(* IEC 61131-3 sources: llm-plc-st-eval/data/definitivo/gemini-3.1-pro-preview/C4/few_shot, 3 files *)

(* ---- ejec_1.st ---- *)
El bloque de función `FB_D` implementa un sistema de control de alternancia y respaldo para dos bombas (sistema de trabajo-reserva o *duty-standby*). Cada vez que se recibe una nueva señal de demanda, el bloque alterna el turno de la bomba principal para garantizar un desgaste uniforme de ambos equipos. Durante la demanda, si la bomba a la que le corresponde el turno presenta una falla, el sistema activa automáticamente la bomba de respaldo y enciende una alarma. Cuando la demanda desaparece, ambas bombas y la alarma se apagan. Esta lógica es ideal para aplicaciones de bombeo de agua, sistemas de presión constante, estaciones de cárcamo, compresores o sistemas de lubricación redundantes donde la fiabilidad y el uso equilibrado de los motores son críticos.

```iecst
FUNCTION_BLOCK FB_D
VAR_INPUT
    demanda : BOOL; (* Señal de peticion de arranque del sistema *)
    falla1 : BOOL;  (* Señal de falla de la bomba 1 *)
    falla2 : BOOL;  (* Señal de falla de la bomba 2 *)
END_VAR
VAR_OUTPUT
    bomba1 : BOOL;   (* Comando de activacion para la bomba 1 *)
    bomba2 : BOOL;   (* Comando de activacion para la bomba 2 *)
    almFalla : BOOL; (* Alarma de falla en la bomba titular del turno *)
END_VAR
VAR
    turno : BOOL;    (* Bandera para alternar el turno (TRUE = Bomba 1, FALSE = Bomba 2) *)
    fDem : R_TRIG;   (* Detector de flanco de subida para la señal de demanda *)
END_VAR

(* Deteccion del flanco de subida de la señal de demanda *)
fDem(CLK := demanda);

(* Alternancia de turno con cada nueva demanda para equilibrar el desgaste *)
IF fDem.Q THEN
    turno := NOT turno;
END_IF

(* Logica de control de bombas mientras exista demanda *)
IF demanda THEN
    IF turno THEN
        (* Turno de la bomba 1 como principal *)
        bomba1 := NOT falla1;            (* Enciende bomba 1 si no tiene falla *)
        bomba2 := falla1 AND NOT falla2; (* Respaldo: enciende bomba 2 si la 1 falla y la 2 esta disponible *)
        almFalla := falla1;              (* Activa alarma si la bomba titular (1) falla *)
    ELSE
        (* Turno de la bomba 2 como principal *)
        bomba2 := NOT falla2;            (* Enciende bomba 2 si no tiene falla *)
        bomba1 := falla2 AND NOT falla1; (* Respaldo: enciende bomba 1 si la 2 falla y la 1 esta disponible *)
        almFalla := falla2;              (* Activa alarma si la bomba titular (2) falla *)
    END_IF
ELSE
    (* Apagado general del sistema cuando no hay demanda *)
    bomba1 := FALSE;
    bomba2 := FALSE;
    almFalla := FALSE;
END_IF
END_FUNCTION_BLOCK
```

(* ---- ejec_2.st ---- *)
Este bloque de función (FB_D) controla un sistema redundante de dos bombas con alternancia automática y lógica de respaldo (failover). Cada vez que se recibe una nueva señal de demanda, el sistema alterna el "turno" de la bomba principal para garantizar un desgaste equitativo entre ambas. Si la bomba a la que le corresponde el turno presenta una falla, el bloque arranca automáticamente la bomba de respaldo (siempre que esta no esté en falla también) y activa una alarma. Cuando la demanda desaparece, ambas bombas y la alarma se apagan. Esta lógica es ideal para aplicaciones de alta disponibilidad como estaciones de bombeo de agua potable, sistemas de achique (cárcamos), o circuitos de refrigeración/calefacción (HVAC) donde se requiere rotación de equipos y seguridad ante fallos.

```iecst
FUNCTION_BLOCK FB_D
VAR_INPUT
    demanda : BOOL; (* Señal de peticion de arranque del sistema *)
    falla1 : BOOL;  (* Señal de falla de la bomba 1 *)
    falla2 : BOOL;  (* Señal de falla de la bomba 2 *)
END_VAR
VAR_OUTPUT
    bomba1 : BOOL;   (* Comando de arranque para la bomba 1 *)
    bomba2 : BOOL;   (* Comando de arranque para la bomba 2 *)
    almFalla : BOOL; (* Alarma de falla de la bomba en turno *)
END_VAR
VAR
    turno : BOOL;    (* Memoria de alternancia (TRUE = Bomba 1, FALSE = Bomba 2) *)
    fDem : R_TRIG;   (* Detector de flanco de subida para la señal de demanda *)
END_VAR

(* Deteccion del flanco de subida de la demanda *)
fDem(CLK := demanda);

(* Alternancia del turno de la bomba principal en cada nueva demanda *)
IF fDem.Q THEN
    turno := NOT turno;
END_IF

(* Logica de control mientras la demanda este activa *)
IF demanda THEN
    IF turno THEN
        (* Turno de la bomba 1 como principal *)
        bomba1 := NOT falla1;                    (* Arranca bomba 1 si no tiene falla *)
        bomba2 := falla1 AND NOT falla2;         (* Respaldo: arranca bomba 2 si la 1 falla y la 2 esta disponible *)
        almFalla := falla1;                      (* Activa alarma si la bomba principal del turno fallo *)
    ELSE
        (* Turno de la bomba 2 como principal *)
        bomba2 := NOT falla2;                    (* Arranca bomba 2 si no tiene falla *)
        bomba1 := falla2 AND NOT falla1;         (* Respaldo: arranca bomba 1 si la 2 falla y la 1 esta disponible *)
        almFalla := falla2;                      (* Activa alarma si la bomba principal del turno fallo *)
    END_IF
ELSE
    (* Si no hay demanda, se apagan las bombas y la alarma *)
    bomba1 := FALSE;
    bomba2 := FALSE;
    almFalla := FALSE;
END_IF
END_FUNCTION_BLOCK
```

(* ---- ejec_3.st ---- *)
Este bloque de función (FB_D) controla un sistema redundante de dos bombas con alternancia automática y respaldo por falla. Cada vez que se recibe una nueva señal de demanda, el sistema alterna el "turno" de la bomba titular para equilibrar el desgaste mecánico de ambos equipos. Durante la operación, si la bomba que tiene el turno presenta una falla, el sistema activa automáticamente la bomba de respaldo (siempre y cuando esta no tenga falla también) y emite una alarma. Cuando no hay demanda, ambas bombas y la alarma se apagan. Es una aplicación clásica y muy útil para estaciones de bombeo de agua, sistemas de achique, circuitos de refrigeración o sistemas de lubricación donde se requiere alta disponibilidad y desgaste uniforme.

```iecst
FUNCTION_BLOCK FB_D
VAR_INPUT
    demanda : BOOL; (* Señal de peticion de arranque del sistema *)
    falla1 : BOOL;  (* Señal de falla de la bomba 1 *)
    falla2 : BOOL;  (* Señal de falla de la bomba 2 *)
END_VAR
VAR_OUTPUT
    bomba1 : BOOL;   (* Comando de arranque para la bomba 1 *)
    bomba2 : BOOL;   (* Comando de arranque para la bomba 2 *)
    almFalla : BOOL; (* Alarma indicadora de falla en la bomba titular *)
END_VAR
VAR
    turno : BOOL;    (* Bandera de alternancia (TRUE = Bomba 1 titular, FALSE = Bomba 2 titular) *)
    fDem : R_TRIG;   (* Detector de flanco de subida para la señal de demanda *)
END_VAR

(* Detecta el instante en que inicia una nueva demanda *)
fDem(CLK := demanda);

(* Alterna el turno de las bombas en cada nuevo arranque para igualar el desgaste *)
IF fDem.Q THEN
    turno := NOT turno;
END_IF

(* Logica de operacion mientras exista demanda *)
IF demanda THEN
    IF turno THEN
        (* --- Turno de la Bomba 1 como titular --- *)
        bomba1 := NOT falla1;                   (* La bomba 1 opera si no tiene falla *)
        bomba2 := falla1 AND NOT falla2;        (* La bomba 2 entra al relevo si la 1 falla y la 2 esta sana *)
        almFalla := falla1;                     (* Se activa la alarma si la bomba titular (1) falla *)
    ELSE
        (* --- Turno de la Bomba 2 como titular --- *)
        bomba2 := NOT falla2;                   (* La bomba 2 opera si no tiene falla *)
        bomba1 := falla2 AND NOT falla1;        (* La bomba 1 entra al relevo si la 2 falla y la 1 esta sana *)
        almFalla := falla2;                     (* Se activa la alarma si la bomba titular (2) falla *)
    END_IF
ELSE
    (* Si no hay demanda, se apagan todos los equipos y la alarma *)
    bomba1 := FALSE;
    bomba2 := FALSE;
    almFalla := FALSE;
END_IF
END_FUNCTION_BLOCK
```
